{region 'Documentation'}
(*!
<summary>Checks whether the REAL value is inside the inclusive range.</summary>
<description>

Minimum &gt; Maximum reports Error during active evaluation; equal bounds are
valid.

All checked operands and bounds must be finite; NaN or either infinity reports Error
during active evaluation.

Numeric diagnostics use the formatter's default six significant digits; rounding affects
the message only, not the comparison.

</description>
*)
{endregion}
FUNCTION_BLOCK AssertInRange_Real EXTENDS AssertionBase
VAR_INPUT
    IN : REAL; //! Actual value checked or observed by this Assertion.
    Minimum : REAL; //! Inclusive lower bound of the comparison; for a range, must not exceed Maximum.
    Maximum : REAL; //! Inclusive upper bound of the comparison; for a range, must not be below Minimum.
END_VAR

SUPER^();

{region 'Documentation'}
(*!
<summary>Check whether the REAL value is inside the inclusive range.</summary>
*)
{endregion}
METHOD PROTECTED Assert
VAR
    Message : STRING(GVL_Constants.MessageLength);
    MinimumText : STRING(GVL_Constants.AssertionValueLength);
    MaximumText : STRING(GVL_Constants.AssertionValueLength);
    ActualText : STRING(GVL_Constants.AssertionValueLength);
END_VAR
IF NOT EvaluationActive THEN
    RETURN;
END_IF;

IF Result = E_Result.Error THEN
    RETURN;
END_IF;

IF NOT Tc2_Utilities.RealIsFinite(x := IN) THEN
    Error(Message := 'Assertion error: IN must be finite.');
    RETURN;
END_IF;

IF NOT Tc2_Utilities.RealIsFinite(x := Minimum) THEN
    Error(Message := 'Assertion error: Minimum must be finite.');
    RETURN;
END_IF;

IF NOT Tc2_Utilities.RealIsFinite(x := Maximum) THEN
    Error(Message := 'Assertion error: Maximum must be finite.');
    RETURN;
END_IF;

IF Minimum > Maximum THEN
    MinimumText := CreateAssertionTextValue_Real(Value := Minimum);
    MaximumText := CreateAssertionTextValue_Real(Value := Maximum);
    Message := CONCAT('Assertion error: minimum exceeds maximum. Minimum = ',
        MinimumText);
    Message := CONCAT(Message, ', Maximum = ');
    Message := CONCAT(Message, MaximumText);
    Message := CONCAT(Message, '.');
    Error(Message := Message);
    RETURN;
END_IF;

IF Result = E_Result.Failed THEN
    RETURN;
END_IF;

IF (IN < Minimum) OR (IN > Maximum) THEN
    MinimumText := CreateAssertionTextValue_Real(Value := Minimum);
    MaximumText := CreateAssertionTextValue_Real(Value := Maximum);
    ActualText := CreateAssertionTextValue_Real(Value := IN);
    Message := CONCAT('Assertion failed: value is outside allowed range. Minimum = ',
        MinimumText);
    Message := CONCAT(Message, ', Maximum = ');
    Message := CONCAT(Message, MaximumText);
    Message := CONCAT(Message, ', Actual = ');
    Message := CONCAT(Message, ActualText);
    Message := CONCAT(Message, '.');
    Fail(Message := Message);
    RETURN;
END_IF;

Pass();
END_METHOD

END_FUNCTION_BLOCK

(* stored: Version 1.1.0.1
   POU AssertInRange_Real: Id {2909fba0-04a1-4491-9e37-6fc335f34379}, SpecialFunc None
   Folder Internal: Id {1fb02e30-7a8e-458a-85f8-94a122ef2b70}
   Method Assert: Id {d56f602c-333b-4395-8d6a-090f40efc20f} *)
